(* IEC 61131-3 sources: SRCI_CLIENT_PLC/RobotLibrary/Library/POUs/ConveyorTracking/MC_SyncToConveyor/Structures, 4 files *)

(* ---- SyncToConveyorOutCmd.st ---- *)
{attribute 'pack_mode' := '1'}
// -------------------------------------------------------------------------
//  SRCI Robot Library
// -------------------------------------------------------------------------
//
//  Object:      SyncToConveyorOutCmd
//  Author:      Thorsten Brach
//  Date:        2024-06-11
//
//  Description:
//
//
//  Copyright:
//    (C) 2024 Thorsten Brach. All rights reserved
//             Licensed under the MIT License.
//
//  Disclaimer:
//    This project is provided without any guarantee and can be used for
//    private and commercial purposes. Any use is at the user’s
//    own risk and responsibility.
//
// -------------------------------------------------------------------------
TYPE SyncToConveyorOutCmd :
STRUCT
  /// Relates to ListenerID >0
  /// Number of successful trigger-based command invocations - For more information refer TO chapter 5.5.12.4
  InvocationCounter      : USINT;
  /// Reserve
  Reserve                : BYTE;
  /// Unique system-generated ID of the "Action" when the function is triggered.
  /// • >0: The "Action" is started by the trigger funcrion with identical FollowID.
  /// • <0: The "Action" is stopped by the trigger function with identical FollowID.
  /// For more information see chapter 5.5.12.4 EmitterID, ListenerID, FollowID and OriginID
  OriginID               : INT;
  /// The TCP is in synchronization with the object on the conveyor belt.
  InSync                 : BOOL;
END_STRUCT
END_TYPE

(* ---- SyncToConveyorParCmd.st ---- *)
{attribute 'pack_mode' := '1'}
// -------------------------------------------------------------------------
//  SRCI Robot Library
// -------------------------------------------------------------------------
//
//  Object:      SyncToConveyorParCmd
//  Author:      Thorsten Brach
//  Date:        2024-06-11
//
//  Description:
//
//
//  Copyright:
//    (C) 2024 Thorsten Brach. All rights reserved
//             Licensed under the MIT License.
//
//  Disclaimer:
//    This project is provided without any guarantee and can be used for
//    private and commercial purposes. Any use is at the user’s
//    own risk and responsibility.
//
// -------------------------------------------------------------------------
TYPE SyncToConveyorParCmd :
STRUCT
  /// Index of assigned conveyor
  ConveyorNo      : USINT;
  /// Define the index number of the UCS that will be assigned to the conveyor.
  /// For more information refer to chapter 5.5.14
  FrameNo         : USINT;
  /// Defines when synchronization starts.
  SyncInMode      : SyncInMode;
  /// Relates to "SyncInMode" "After distance" (1) and "After time" (2):
  /// Parameter for the synchronization
  /// • "After distance" (1)
  ///    •  Distance in mm
  /// • "After time" (2)
  ////   • Time in ms
  SyncInParameter : REAL;
  /// Define the maximum adjustment velocity for the robot to catch up to the conveyor belt.
  /// The velocity must be greater than the velocity of the conveyor belt.
  /// • 0 (default): no limit
  ///       o No conveyor tracking specific limit
  ///       o RC internal limit applies
  /// • >0: use limit
  ///       o Conveyor tracking specific limit applies
  MaxVelocity     : REAL;
  /// Define the maximum adjustment acceleration for the robot to catch up to the conveyor belt.
  /// • 0 (default): no limit
  ///     o No conveyor tracking specific limit
  ///     o RC internal limit applies
  /// • >0: use limit
  ///     o Conveyor tracking specific limit applies
  MaxAcceleration : REAL;
  /// ID of associated trigger function:
  ///  •  0: No Trigger (default):
  ///        o No trigger related behavior
  ///  • >0: Trigger:
  ///        o Start executing, when the trigger function with the identical EmitterID is triggered.
  /// Always positive.
  /// For more information, see chapter 5.5.12 Triggers
  ListenerID      : SINT;
END_STRUCT
END_TYPE

(* ---- SyncToConveyorRecvData.st ---- *)
{attribute 'pack_mode' := '1'}
// -------------------------------------------------------------------------
//  SRCI Robot Library
// -------------------------------------------------------------------------
//
//  Object:      SyncToConveyorRecvData
//  Author:      Thorsten Brach
//  Date:        2024-06-11
//
//  Description:
//
//
//  Copyright:
//    (C) 2024 Thorsten Brach. All rights reserved
//             Licensed under the MIT License.
//
//  Disclaimer:
//    This project is provided without any guarantee and can be used for
//    private and commercial purposes. Any use is at the user’s
//    own risk and responsibility.
//
// -------------------------------------------------------------------------
TYPE SyncToConveyorRecvData EXTENDS RspHeader :
STRUCT
  InvocationCounter : USINT;
  /// Reserve
  Reserved          : SINT;
  /// Unique system-generated ID of the "Action" when the function is triggered.
  /// • >0: The "Action" is started by the trigger funcrion with identical FollowID.
  /// • <0: The "Action" is stopped by the trigger function with identical FollowID.
  /// For more information see chapter 5.5.12.4 EmitterID, ListenerID, FollowID and OriginID
  OriginID          : INT;
  /// The TCP is in synchronization with the object on the conveyor belt.
  InSync            : BOOL;
END_STRUCT
END_TYPE

(* ---- SyncToConveyorSendData.st ---- *)
{attribute 'pack_mode' := '1'}
// -------------------------------------------------------------------------
//  SRCI Robot Library
// -------------------------------------------------------------------------
//
//  Object:      SyncToConveyorSendData
//  Author:      Thorsten Brach
//  Date:        2024-06-11
//
//  Description:
//
//
//  Copyright:
//    (C) 2024 Thorsten Brach. All rights reserved
//             Licensed under the MIT License.
//
//  Disclaimer:
//    This project is provided without any guarantee and can be used for
//    private and commercial purposes. Any use is at the user’s
//    own risk and responsibility.
//
// -------------------------------------------------------------------------
TYPE SyncToConveyorSendData EXTENDS CmdHeader:
STRUCT
  /// EmitterID
  EmitterID       : ARRAY[0..3] OF SINT;
  /// ID of associated trigger function:
  /// • 0: No Trigger (default): No trigger related behavior
  /// • >0: Trigger: o Start executing, when the trigger function with the identical EmitterID is triggered.
  /// Always positive.
  /// For more information, see chapter 5.5.12 Triggers
  ListenerID      : SINT;
  /// Reserve
  Reserve         : BYTE;
  /// Index of assigned conveyor
  ConveyorNo      : USINT;
  /// Define the index number of the UCS that will be assigned to the conveyor.
  /// For more information refer to chapter 5.5.14
  FrameNo         : USINT;
  /// Defines when synchronization starts
  SyncInMode      : SyncInMode;
  /// Relates to "SyncInMode" "After distance" (1) and "After time" (2): Parameter for the synchronization
  /// • "After distance" (1) -  Distance in mm
  /// • "After time" (2) -  Time in ms
  SyncInParameter : REAL;
  /// Define the maximum adjustment velocity for the robot to catch up to the conveyor belt.
  /// The velocity must be greater than the velocity of the conveyor belt.
  /// • 0 (default): no limit - No conveyor tracking specific limit
  ///                         - RC internal limit applies
  /// • >0: use limit         - Conveyor tracking specific limit applies
  MaxVelocity     : REAL;
  /// Define the maximum adjustment acceleration for the robot to catch up to the conveyor belt.
  /// • 0 (default): no limit - No conveyor tracking specific limit
  ///                         - RC internal limit applies
  /// • >0: use limit         - Conveyor tracking specific limit applies
  MaxAcceleration : REAL;
  /// ID of associated trigger function:
  /// • 0: No Trigger (default): No trigger related behavior
  /// • >0: Trigger:  Start executing, when the trigger function with the identical EmitterID is triggered.
  /// Always positive.
  /// For more information, see chapter 5.5.12 Triggers
END_STRUCT
END_TYPE
